FUNCTION_BLOCK FB_Blocks
VAR
    nA, nB, nSum, nCopy : INT;
    bHigh : BOOL;
END_VAR
VAR // added by the converter: edge detectors and wires of the graphical bodies
    _w1 : INT;
END_VAR

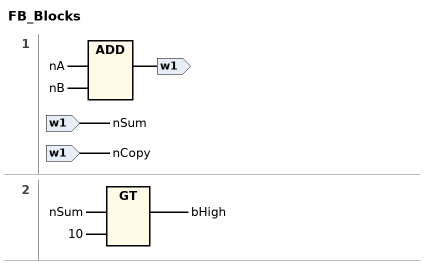
// NETWORK 1
_w1 := nA + nB;
nSum := _w1;
nCopy := _w1;

// NETWORK 2
bHigh := nSum > 10;

END_FUNCTION_BLOCK

(* stored: Version 1.1.0.1, ProductVersion 3.1.4024.12
   POU FB_Blocks: Id {00000000-0000-0000-0000-000000000001}, SpecialFunc None *)
